Fanuc KAREL source: KA00152.KL

PROGRAM KA00152
%NOLOCKGROUP
VAR
  SRC: ARRAY[4] OF INTEGER
  DST: ARRAY[4] OF XYZWPR
BEGIN
  DST = SRC
END KA00152
